Fanuc KAREL source: KB00148.KL

PROGRAM KB00148
%NOLOCKGROUP
%ENVIRONMENT MEMO
VAR
  P1: STRING[80]
  P2: STRING[80]
  P3: INTEGER
BEGIN
  P1 = 'A'
  P2 = 'A'
  P3 = 1
  RENAME_VARS(P1, P2, P3)
END KB00148
